(* IEC 61131-3 sources: IRIS-Project/LASAL CONTROL SOFTWARE/LasalProject_2025_09_12/Runtime/%LASALAPPDATA%/Runtime/Library/Loader/Class/MMServerBase, 1 file *)

(* ---- MMServerBase.st ---- *)
#pragma warning(disable:73);

FUNCTION VIRTUAL GLOBAL MMServerBase::WriteDataOff
	VAR_INPUT
		udLen 	: UDINT;
		udOff 	: UDINT;
		pData 	: ^USINT;
	END_VAR

END_FUNCTION

FUNCTION VIRTUAL GLOBAL MMServerBase::GetCharSize
	VAR_INPUT
		nBufferId 	: UDINT;
	END_VAR
	VAR_OUTPUT
		usSize 	: USINT;
	END_VAR

  usSize := 0;

END_FUNCTION

FUNCTION VIRTUAL GLOBAL MMServerBase::GetCRC
	VAR_OUTPUT
		udCRC 	: UDINT;
	END_VAR

  udCRC := 0;

END_FUNCTION

FUNCTION VIRTUAL GLOBAL MMServerBase::GetDataAt
	VAR_INPUT
		pData 	: ^USINT;
		udSize 	: UDINT;
		udAt 	: UDINT;
	END_VAR

END_FUNCTION

FUNCTION VIRTUAL GLOBAL MMServerBase::GetBufferLen
	VAR_INPUT
		nBufferId 	: UDINT;
	END_VAR
	VAR_OUTPUT
		udLen 	: UDINT;
	END_VAR

  udLen:= 0;

END_FUNCTION

FUNCTION VIRTUAL GLOBAL MMServerBase::ReadDataOff
	VAR_INPUT
		udOff 	: UDINT;
		pData 	: ^USINT;
		udMax 	: UDINT;
	END_VAR
	VAR_OUTPUT
		udLen 	: UDINT;
	END_VAR

  udLen := 0;

END_FUNCTION

FUNCTION VIRTUAL GLOBAL MMServerBase::GetDataPtrIn
	VAR_OUTPUT
		pData 	: ^USINT;
	END_VAR

  pData := NIL;

END_FUNCTION

#pragma warning(default:73);
